(* IEC 61131-3 sources: kns-port-domestic/targets/astra/lib/src/DUTs/AnalogInput, 8 files *)

(* ---- E_AiAlarm.dut.st ---- *)
// Назначение: индексы слотов тревог аналогового входа (afbAlarm[i], astAlarm[i]) и уставок
//             (astLimit[HH..LL]). Нестрогое перечисление: им индексируются массивы.
// Автор:      kr0nsch
// Версия:     0.1.0
// Документ:   docs/fb/FB_AnalogInput.md
{attribute 'qualified_only'}
TYPE E_AiAlarm :
(
    HH         := 0,   // верхняя аварийная уставка
    H          := 1,   // верхняя предупредительная уставка
    L          := 2,   // нижняя предупредительная уставка
    LL         := 3,   // нижняя аварийная уставка
    Failure    := 4,   // подтверждённый отказ сигнала
    OutOfRange := 5    // сигнал вне диапазона измерения (NE 43)
) UINT;
END_TYPE

(* ---- E_AiFailValue.dut.st ---- *)
// Назначение: значение аналогового входа при подтверждённом отказе сигнала.
// Автор:      kr0nsch
// Версия:     0.1.0
// Документ:   docs/fb/FB_AnalogInput.md
{attribute 'qualified_only'}
{attribute 'strict'}
TYPE E_AiFailValue :
(
    HoldLast   := 0,   // удерживать последнее хорошее значение
    Substitute := 1    // подставить stCfg.rFailValue_eu
) INT;
END_TYPE

(* ---- E_AiInputType.dut.st ---- *)
// Назначение: смысл входа rIn аналогового входа и применимость проверки NAMUR NE 43.
// Автор:      kr0nsch
// Версия:     0.1.0
// Документ:   docs/fb/FB_AnalogInput.md
{attribute 'qualified_only'}
{attribute 'strict'}
TYPE E_AiInputType :
(
    MilliAmp := 0,   // rIn в мА, 4–20, проверка NE 43
    Norm420  := 1,   // rIn 0..1 соответствует 4–20 мА; NE 43 по пересчёту I = 4 + 16·rIn
    Norm01   := 2,   // rIn 0..1 без NE 43 (0–10 В и т. п.)
    Eng      := 3,   // rIn уже в инж. ед. (Modbus REAL, расчёт); NE 43 не применяется
    Raw      := 4    // rIn в единицах канала (отсчёты АЦП, целое из Modbus): rRawLo_cnt..rRawHi_cnt
) INT;
END_TYPE

(* ---- E_AiSignalState.dut.st ---- *)
// Назначение: мгновенная классификация сигнала аналогового входа (до задержки
//             подтверждения). Границы NE 43 — сверить с NAMUR NE 43 (A-02).
// Автор:      kr0nsch
// Версия:     0.1.0
// Документ:   docs/fb/FB_AnalogInput.md
{attribute 'qualified_only'}
{attribute 'strict'}
TYPE E_AiSignalState :
(
    Good         := 0,
    UnderRange   := 1,   // 3,6 < I < 3,8 мА
    OverRange    := 2,   // 20,5 < I < 21,0 мА
    FailLow      := 3,   // I <= 3,6 мА
    FailHigh     := 4,   // I >= 21,0 мА
    ChannelFault := 5,   // xChannelFault
    NotFinite    := 6    // NaN, ±Inf, |rIn| > REAL_SANE_MAX
) INT;
END_TYPE

(* ---- ST_AiLimitCfg.dut.st ---- *)
// Назначение: параметры одной уставки (FB_LimitMonitor, astLimit[i] аналогового входа).
//             Тип лежит в Persistent Variables приложения и заморожен в пределах 1.x (A-13).
// Автор:      kr0nsch
// Версия:     0.1.0
// Документ:   docs/fb/FB_LimitMonitor.md
{attribute 'qualified_only'}
TYPE ST_AiLimitCfg :
STRUCT
    xEnable      : BOOL := FALSE;   // уставка включена
    rSetpoint_eu : REAL := 0.0;     // уставка, инж. ед.
    rHyst_eu     : REAL := 0.0;     // гистерезис, инж. ед., >= 0
    tOnDelay     : TIME := T#0S;    // задержка срабатывания флага
    tOffDelay    : TIME := T#0S;    // задержка снятия флага
END_STRUCT
END_TYPE

(* ---- ST_AnalogInputCfg.dut.st ---- *)
// Назначение: параметры аналогового входа (Persistent Variables приложения,
//             VAR_IN_OUT CONSTANT stCfg). Значения по умолчанию проходят CheckConfig.
//             Тип лежит в Persistent Variables приложения и заморожен в пределах 1.x (A-13).
// Автор:      kr0nsch
// Версия:     0.1.0
// Документ:   docs/fb/FB_AnalogInput.md
{attribute 'qualified_only'}
TYPE ST_AnalogInputCfg :
STRUCT
    eInput         : E_AiInputType := E_AiInputType.MilliAmp;
    rRangeLo_eu    : REAL := 0.0;      // значение при 4 мА / 0.0
    rRangeHi_eu    : REAL := 100.0;    // значение при 20 мА / 1.0 / rRawHi_cnt
    rRawLo_cnt     : REAL := 0.0;      // только Raw: значение канала, соответствующее rRangeLo_eu
    rRawHi_cnt     : REAL := 0.0;      // только Raw: значение канала, соответствующее rRangeHi_eu (0/0 — не задано)
    xSqrt          : BOOL := FALSE;    // корень (расход по перепаду давления)
    rLowCut_pct    : REAL := 0.0;      // отсечка малых значений, % шкалы (после корня); 0 — нет
    tFilter        : TIME := T#0S;     // постоянная времени фильтра; T#0S — без фильтра
    tFailDelay     : TIME := T#2S;     // подтверждение отказа / выхода за диапазон и возврата
    eFailValue     : E_AiFailValue := E_AiFailValue.HoldLast;
    rFailValue_eu  : REAL := 0.0;      // значение при Substitute
    xLimitsOnFail  : BOOL := FALSE;    // TRUE — при подтверждённом отказе уставки считаются по значению отказа
    xClamp         : BOOL := FALSE;    // ограничить значение шкалой (по умолчанию — экстраполяция)
    astLimit       : ARRAY[0..3] OF ST_AiLimitCfg;   // индекс E_AiAlarm.HH, H, L, LL
    tSubstMax      : TIME := T#8H;     // макс. длительность подмены; T#0S — без ограничения
    udiAlarmIdBase : UDINT := 0;       // номер первой тревоги устройства (dev_no * 10)
    astAlarm       : ARRAY[0..GVL_Const.DEV_ALARMS_MAX - 1] OF ST_AlarmCfg := [
        (ePriority := E_AlarmPriority.High),      // 0 HH
        (ePriority := E_AlarmPriority.Low),       // 1 H
        (ePriority := E_AlarmPriority.Low),       // 2 L
        (ePriority := E_AlarmPriority.High),      // 3 LL
        (ePriority := E_AlarmPriority.Medium),    // 4 Failure
        (ePriority := E_AlarmPriority.Low),       // 5 OutOfRange
        (ePriority := E_AlarmPriority.None),      // 6 —
        (ePriority := E_AlarmPriority.None)];     // 7 —
END_STRUCT
END_TYPE

(* ---- ST_AnalogInputCmd.dut.st ---- *)
// Назначение: команды HMI/SCADA аналогового входа (GVL_Hmi приложения, VAR_IN_OUT stCmd).
// Автор:      kr0nsch
// Версия:     0.1.0
// Документ:   docs/fb/FB_AnalogInput.md
{attribute 'qualified_only'}
TYPE ST_AnalogInputCmd :
STRUCT
    stCommon       : ST_DeviceCmd;   // xSetAuto — «Измерение», xSetManual — «Подмена», xSetOos
    rSubstValue_eu : REAL;           // значение подмены; в Auto ФБ пишет сюда текущее rValue_eu
END_STRUCT
END_TYPE

(* ---- ST_AnalogInputSts.dut.st ---- *)
// Назначение: состояние аналогового входа для HMI/SCADA. 44 байта, 22 регистра Modbus:
//             только 16- и 32-битные поля без скрытого выравнивания.
// Автор:      kr0nsch
// Версия:     0.1.0
// Документ:   docs/fb/FB_AnalogInput.md
{attribute 'qualified_only'}
TYPE ST_AnalogInputSts :
STRUCT
    stCommon        : ST_DeviceSts;      // 0..27
    rValue_eu       : REAL;              // 28: итоговое значение
    rValue_pct      : REAL;              // 32: % шкалы
    rIn             : REAL;              // 36: сырое значение входа
    eSignal         : E_AiSignalState;   // 40: мгновенная классификация (до задержки)
    uiSubstRemain_s : UINT;              // 42: до автоматического снятия подмены, с; 0 — подмены нет
END_STRUCT
END_TYPE
